INTERFACE I_Cooling

PROPERTY bRunning : BOOL
GET
END_GET
END_PROPERTY

PROPERTY nSpeed : REAL
GET
END_GET
END_PROPERTY

END_INTERFACE

(* stored: Version 1.1.0.1
   Itf I_Cooling: Id {7df69075-8e3e-46a8-bee5-ca7f72ad12ae}
   Property bRunning: Id {43ef9597-4711-4a66-b9c0-3a23e97fcd2d}
   Get Get: Id {dceadee5-c63a-435b-a1ca-8eb738453e10}
   Property nSpeed: Id {0dcdc53e-d53a-4e05-83b7-56423b4ce12d}
   Get Get: Id {b74fe025-7dbc-4236-8385-6f1164e9c003} *)
